FUNCTION_BLOCK IO_RouteAO (* Picks the way an IO block reaches its signal from the Address (a Pi line, a local IO handle, Modbus or simulated) and passes values through that way only. Technical: Backend router for IO_AO; Address: 'gpio[chip:line(:pull_up|:pull_down)(:active_low)]' or 'pwm[chip:channel:period_ns]' a Raspberry Pi's line, set up here; 'modbus[...]' a Modbus CLIENT ID; 'sim' simulated; another name a local IO handle set up elsewhere (IX/QX PARAMS); empty: not connected (QO = FALSE) *)
  (* Standard: 61499-2 *)
  (* Version 0.1, 2026-09-28, Project contributors, AAU Smart Production Lab *)
  PACKAGE modlib;
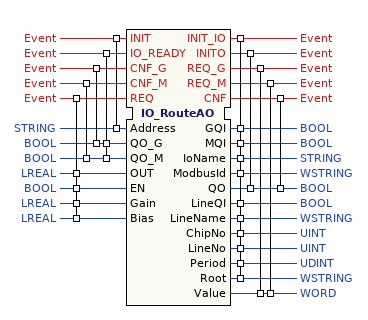
  EVENT_INPUT
    INIT WITH Address; (* Work out from Address how the point is reached *)
    IO_READY WITH QO_G, QO_M; (* The line, the local IO block and the Modbus client are initialised *)
    CNF_G WITH QO_G; (* The local IO block answered *)
    CNF_M WITH QO_M; (* The Modbus client answered *)
    REQ WITH OUT, EN, Gain, Bias; (* Access the point *)
  END_EVENT
  EVENT_OUTPUT
    INIT_IO WITH GQI, MQI, IoName, ModbusId, LineQI, LineName, ChipNo, LineNo, Period, Root; (* Set up the line, the local IO block and the Modbus client (each only if it is the way) *)
    INITO WITH QO; (* Initialised: QO says whether the point is reachable *)
    REQ_G WITH Value; (* Access the point through the local IO block (IX/QX/IW/QW) *)
    REQ_M WITH Value; (* Access the point through the Modbus client *)
    CNF WITH QO; (* Done: QO says whether it worked *)
  END_EVENT
  VAR_INPUT
    Address : STRING; (* Where the point is: 'gpio[chip:line(:pull_up|:pull_down)(:active_low)]', 'pwm[chip:channel:period_ns]', 'modbus[...]', 'sim', or an IO handle's name; empty: not connected *)
    QO_G : BOOL; (* The local IO block works *)
    QO_M : BOOL; (* The Modbus client works *)
    OUT : LREAL; (* The value to write *)
    EN : BOOL; (* On; FALSE writes 0 (no pulses on a PWM channel) *)
    Gain : LREAL := 1.0; (* Raw = Bias + OUT * Gain, limited to 0..65535 *)
    Bias : LREAL; (* Raw = Bias + OUT * Gain, limited to 0..65535 *)
  END_VAR
  VAR_OUTPUT
    GQI : BOOL; (* Use the local IO block *)
    MQI : BOOL; (* Use the Modbus client *)
    IoName : STRING; (* The local IO handle's name (PARAMS of IX/QX/IW/QW) *)
    ModbusId : WSTRING; (* The Modbus CLIENT's ID *)
    QO : BOOL; (* The point is reachable, the last access worked *)
    LineQI : BOOL; (* Set up a Raspberry Pi line here (a gpio[...] or pwm[...] address) *)
    LineName : WSTRING; (* The name the line is registered under (the address) *)
    ChipNo : UINT; (* The GPIO or PWM chip's number *)
    LineNo : UINT; (* The GPIO line's or PWM channel's number *)
    Period : UDINT; (* The PWM period in ns *)
    Root : WSTRING; (* The sysfs PWM folder (empty: /sys/class/pwm) *)
    Value : WORD; (* The raw value to write (0 to 65535 for an analog output) *)
  END_VAR
  VAR
    Backend : USINT;
    Raw : LREAL;
  END_VAR
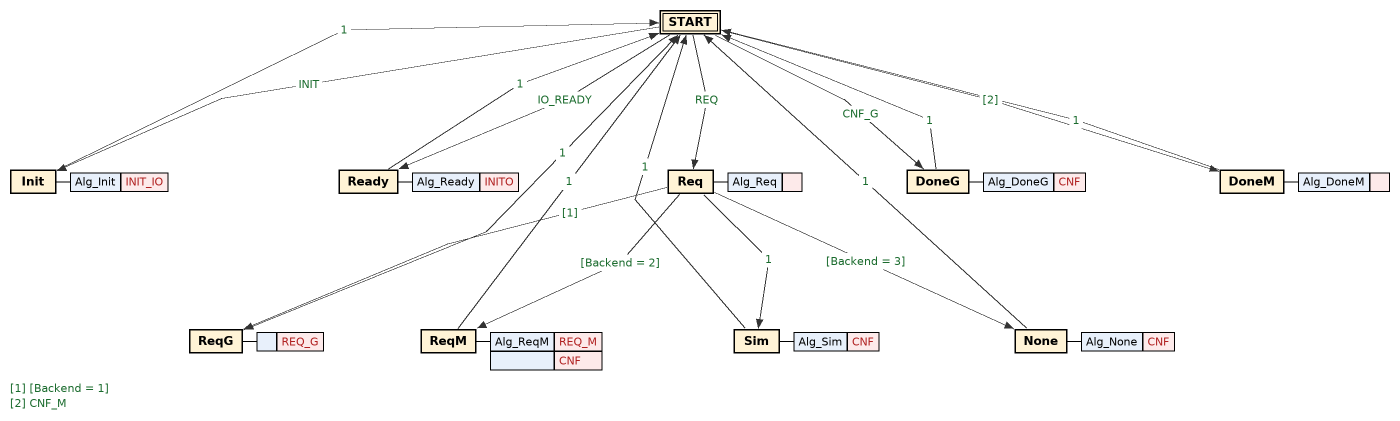
  EC_STATES
    START;
    Init : Alg_Init -> INIT_IO;
    Ready : Alg_Ready -> INITO;
    ReqG : -> REQ_G;
    ReqM : Alg_ReqM -> REQ_M, -> CNF;
    Req : Alg_Req;
    Sim : Alg_Sim -> CNF;
    None : Alg_None -> CNF;
    DoneG : Alg_DoneG -> CNF;
    DoneM : Alg_DoneM;
  END_STATES
  EC_TRANSITIONS
    START TO Init := INIT;
    Init TO START := 1;
    START TO Ready := IO_READY;
    Ready TO START := 1;
    START TO Req := REQ;
    Req TO ReqG := [Backend = 1];
    Req TO ReqM := [Backend = 2];
    Req TO None := [Backend = 3];
    Req TO Sim := 1;
    START TO DoneG := CNF_G;
    START TO DoneM := CNF_M;
    ReqG TO START := 1;
    ReqM TO START := 1;
    Sim TO START := 1;
    None TO START := 1;
    DoneG TO START := 1;
    DoneM TO START := 1;
  END_TRANSITIONS
  ALGORITHM Alg_Init IN ST:
VAR_TEMP
  Field : STRING;
  Length : INT;
  Cut : INT;
  Pos : INT;
  Digit : INT;
  Number : UDINT;
END_VAR
Backend := 3;
LineQI := FALSE;
IF Address = 'sim' THEN
  Backend := 0;
ELSIF LEFT(Address, 7) = 'modbus[' THEN
  Backend := 2;
  ModbusId := STRING_TO_WSTRING(Address);
ELSIF LEFT(Address, 4) = 'pwm[' THEN
  Backend := 1;
  IoName := Address;
  LineQI := TRUE;
  LineName := STRING_TO_WSTRING(Address);
  Length := LEN(Address);
  Field := MID(Address, Length - 4, 5);
  Cut := FIND(Field, ':');
  IF Cut = 0 THEN
    Cut := FIND(Field, ']');
  END_IF;
  Number := 0;
  FOR Digit := 1 TO Cut - 1 DO
    Pos := FIND('0123456789', MID(Field, 1, Digit));
    Number := Number * 10 + INT_TO_UDINT(Pos - 1);
  END_FOR;
  ChipNo := UDINT_TO_UINT(Number);
  Length := LEN(Field);
  Field := MID(Field, Length - Cut, Cut + 1);
  Cut := FIND(Field, ':');
  IF Cut = 0 THEN
    Cut := FIND(Field, ']');
  END_IF;
  Number := 0;
  FOR Digit := 1 TO Cut - 1 DO
    Pos := FIND('0123456789', MID(Field, 1, Digit));
    Number := Number * 10 + INT_TO_UDINT(Pos - 1);
  END_FOR;
  LineNo := UDINT_TO_UINT(Number);
  Length := LEN(Field);
  Field := MID(Field, Length - Cut, Cut + 1);
  Cut := FIND(Field, ':');
  IF Cut = 0 THEN
    Cut := FIND(Field, ']');
  END_IF;
  Number := 0;
  FOR Digit := 1 TO Cut - 1 DO
    Pos := FIND('0123456789', MID(Field, 1, Digit));
    Number := Number * 10 + INT_TO_UDINT(Pos - 1);
  END_FOR;
  Period := (Number);
  Length := LEN(Field);
  Field := MID(Field, Length - Cut, Cut + 1);
  Length := LEN(Field);
  IF Length > 0 THEN
    Root := STRING_TO_WSTRING(LEFT(Field, Length - 1));
  END_IF;
ELSIF LEN(Address) > 0 THEN
  Backend := 1;
  IoName := Address;
END_IF;
GQI := Backend = 1;
MQI := Backend = 2;
  END_ALGORITHM
  ALGORITHM Alg_Ready IN ST:
QO := (Backend = 0) OR ((Backend = 1) AND QO_G) OR ((Backend = 2) AND QO_M);
  END_ALGORITHM
  ALGORITHM Alg_ReqM IN ST:
QO := QO_M;
  END_ALGORITHM
  ALGORITHM Alg_Req IN ST:
IF EN THEN
  Raw := Bias + OUT * Gain;
  IF Raw < 0.0 THEN
    Raw := 0.0;
  ELSIF Raw > 65535.0 THEN
    Raw := 65535.0;
  END_IF;
  Value := UINT_TO_WORD(LREAL_TO_UINT(Raw));
ELSE
  Value := WORD#0;
END_IF;
  END_ALGORITHM
  ALGORITHM Alg_Sim IN ST:
QO := TRUE;
  END_ALGORITHM
  ALGORITHM Alg_None IN ST:
QO := FALSE;
  END_ALGORITHM
  ALGORITHM Alg_DoneG IN ST:
QO := QO_G;
  END_ALGORITHM
  ALGORITHM Alg_DoneM IN ST:
QO := QO_M;
  END_ALGORITHM
END_FUNCTION_BLOCK
